# B&R Automation Studio project lab1
Automation Studio 4.12.10.39

## Configuration Config1

CPU 4PP065.0571-P74, AutomationRuntime D4.52, Build 4.1.2, Vc V4.52.0

### Task classes (Cpu.sw)
```
Cyclic#3:
  Program <- Program.prg
Binaries: udbdef, TCData, iomap, ashwac, Role, sysconf, arconfig, asfw, User, ashwd
Libraries: Library
```

### Hardware
```
4PP065_0571_P74 : 4PP065.0571-P74 v1.2.0.0
  Connector IF4:
    DNAConfiguration = manual
  Connector IF5:
    ActivateDevice = 1
    Mode = Manual
    InternetAddress = 10.0.1.10
    SubnetMask = 255.255.255.0
  ConfigurationID = labBR
  Simulation = 1
```

- Physical/Config1/4PP065_0571_P74/IoMap.iom: same as Physical/Config1/4PP065_0571_P74/Cpu.per
- Physical/Config1/4PP065_0571_P74/PvMap.vvm: same as Physical/Config1/4PP065_0571_P74/Cpu.per
## Logical view

Binary libraries used (declarations not repeated): operator, runtime, astime, AsIecCon


### Program Logical/Program (ANSIC)

#### Cyclic.c - Cyclic code
```c
#include <bur/plctypes.h>

#ifdef _DEFAULT_INCLUDES
#include <AsDefault.h>
#endif

void _CYCLIC ProgramCyclic(void)
{
	/* Cyclic #4 and the model use dt = 2 ms.  This produces a repeating
	   4 s test signal: 1 s at zero, 2 s at 60 rpm, 1 s at zero. */
	if (!Enable) {
		counter=0;
		Speed=0.0;

		return;
	}
	counter++;
	if ((counter >= 400) && (counter < 800))
		Speed=60.0;
	else
		Speed=0.0;

	if (counter >= 800)
		counter=0;

	if (Enable) {
		fb_controller.e=Speed-fb_motor.w;
		FB_Regulator(&fb_controller);
		fb_motor.u=fb_controller.u;
	}
	else {
		fb_motor.u=0.0;
	}

	FB_Motor(&fb_motor);
	fb_motor_2.u=Speed * fb_motor_2.ke;
	FB_Motor(&fb_motor_2);
}
```

#### Init.c - Initialization code
```c
#include <bur/plctypes.h>

#ifdef _DEFAULT_INCLUDES
	#include <AsDefault.h>
#endif

void _INIT ProgramInit(void)
{
	fb_motor.ke=0.00096;
	fb_motor.Tm=0.04;
	fb_motor.dt=0.002;
	fb_motor.w=0.0;
	fb_motor.phi=0.0;
	fb_motor.integrator.out=0.0;

	fb_motor_2.ke=0.00096;
	fb_motor_2.Tm=0.04;
	fb_motor_2.dt=0.002;
	fb_motor_2.w=0.0;
	fb_motor_2.phi=0.0;
	fb_motor_2.integrator.out=0.0;

	fb_controller.k_p=0.000192;
	fb_controller.k_i=0.0048;
	fb_controller.max_abs_value=24.0;
	fb_controller.dt=0.002;
	fb_controller.u=0.0;
	fb_controller.iyOld=0.0;
	fb_controller.integrator.out=0.0;

	Enable=0;
	Speed=0.0;
	counter=0;
}
```

#### Exit.c - Exit code
```c
#include <bur/plctypes.h>

#ifdef _DEFAULT_INCLUDES
	#include <AsDefault.h>
#endif

void _EXIT ProgramExit(void)
{

}
```

#### Variables.var - Local variables
```iecst
VAR
	fb_controller : FB_Regulator;
	fb_motor : FB_Motor;
	fb_motor_2 : FB_Motor;
	Speed : REAL;
	Enable : BOOL;
	counter : UDINT;
END_VAR
```

### Library Logical/Library (ANSIC)

#### Library.fun - Exported functions and function blocks
```iecst
{REDUND_ERROR} {REDUND_UNREPLICABLE} FUNCTION_BLOCK FB_Integrator (*TODO: Add your comment here*) (*$GROUP=User,$CAT=User,$GROUPICON=User.png,$CATICON=User.png*)
	VAR_INPUT
		in : {REDUND_UNREPLICABLE} REAL;
	END_VAR
	VAR_OUTPUT
		out : {REDUND_UNREPLICABLE} REAL;
	END_VAR
	VAR
		dt : {REDUND_UNREPLICABLE} REAL;
	END_VAR
END_FUNCTION_BLOCK

{REDUND_ERROR} {REDUND_UNREPLICABLE} FUNCTION_BLOCK FB_Motor (*TODO: Add your comment here*) (*$GROUP=User,$CAT=User,$GROUPICON=User.png,$CATICON=User.png*)
	VAR_INPUT
		u : {REDUND_UNREPLICABLE} REAL;
	END_VAR
	VAR_OUTPUT
		w : {REDUND_UNREPLICABLE} REAL;
		phi : {REDUND_UNREPLICABLE} REAL;
	END_VAR
	VAR
		integrator : {REDUND_UNREPLICABLE} FB_Integrator;
		Tm : {REDUND_UNREPLICABLE} REAL;
		ke : {REDUND_UNREPLICABLE} REAL;
		dt : {REDUND_UNREPLICABLE} REAL;
	END_VAR
END_FUNCTION_BLOCK

{REDUND_ERROR} {REDUND_UNREPLICABLE} FUNCTION_BLOCK FB_Regulator (*TODO: Add your comment here*) (*$GROUP=User,$CAT=User,$GROUPICON=User.png,$CATICON=User.png*)
	VAR_INPUT
		e : {REDUND_UNREPLICABLE} REAL;
	END_VAR
	VAR_OUTPUT
		u : {REDUND_UNREPLICABLE} REAL;
	END_VAR
	VAR
		k_p : {REDUND_UNREPLICABLE} REAL;
		k_i : {REDUND_UNREPLICABLE} REAL;
		integrator : {REDUND_UNREPLICABLE} FB_Integrator;
		iyOld : {REDUND_UNREPLICABLE} REAL;
		max_abs_value : {REDUND_UNREPLICABLE} REAL;
		dt : {REDUND_UNREPLICABLE} REAL;
	END_VAR
END_FUNCTION_BLOCK
```

#### FB_Integrator.c
```c
#include <bur/plctypes.h>
#ifdef __cplusplus
	extern "C"
	{
#endif
	#include "Library.h"
#ifdef __cplusplus
	};
#endif
/* TODO: Add your comment here */
void FB_Integrator(struct FB_Integrator* inst)
{
	inst->out= inst->out + inst->in * inst->dt;
}
```

#### FB_Motor.c
```c
#include <bur/plctypes.h>
#ifdef __cplusplus
	extern "C"
	{
#endif
	#include "Library.h"
#ifdef __cplusplus
	};
#endif
/* TODO: Add your comment here */
void FB_Motor(struct FB_Motor* inst)
{
	REAL e;

	e=inst->u/inst->ke-inst->w;
	inst->integrator.in=e/inst->Tm;
	inst->integrator.dt=inst->dt;
	FB_Integrator(&inst->integrator);

	inst->w= inst->integrator.out;
	/* w is measured in rpm, while phi is measured in radians. */
	inst->phi=inst->phi + inst->w * 0.1047197551 * inst->dt;
}
```

#### FB_Regulator.c
```c
#include <bur/plctypes.h>

#ifdef __cplusplus
extern "C"
{
#endif
#include "Library.h"
#ifdef __cplusplus
};
#endif

void FB_Regulator(struct FB_Regulator* inst)
{
	REAL p_term;
	REAL sum_before_sat;
	REAL u_sat;

	/* Пропорциональная составляющая */
	p_term=inst->e * inst->k_p;

	/* Ограничитель после П-звена */
	if (p_term > inst->max_abs_value)
		p_term=inst->max_abs_value;
	else if (p_term < -inst->max_abs_value)
		p_term=-inst->max_abs_value;

	/* Интегратор с предыдущей поправкой противонакопления */
	inst->integrator.in=
		inst->e * inst->k_i + inst->iyOld;

	inst->integrator.dt=inst->dt;
	FB_Integrator(&inst->integrator);

	/* Неограниченный выход ПИ-регулятора */
	sum_before_sat=p_term + inst->integrator.out;

	/* Ограничитель выходного напряжения */
	if (sum_before_sat > inst->max_abs_value)
		u_sat=inst->max_abs_value;
	else if (sum_before_sat < -inst->max_abs_value)
		u_sat=-inst->max_abs_value;
	else
		u_sat=sum_before_sat;

	/* Сохраняем именно поправку противонакопления */
	inst->iyOld=u_sat-sum_before_sat;
	inst->u=u_sat;
}
```
